(* CoDeSys 2.3 export: ld.exp *)

(* POU PLC_LD_PRG_TR, LD *)
PROGRAM PLC_LD_PRG_TR
VAR
END_VAR
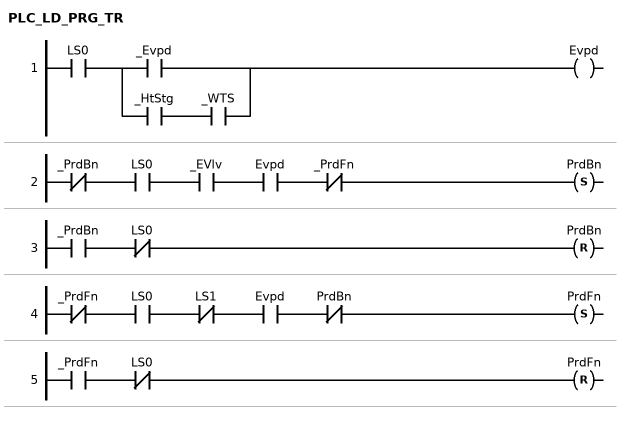
_LD_ (* Ladder Diagram *)
NETWORK 1
	[LS0] - { [_Evpd] | [_HtStg] - [_WTS] } --- (Evpd)
NETWORK 2
	[/_PrdBn] - [LS0] - [_EVlv] - [Evpd] - [/_PrdFn] --- (S PrdBn)
NETWORK 3
	[_PrdBn] - [/LS0] --- (R PrdBn)
NETWORK 4
	[/_PrdFn] - [LS0] - [/LS1] - [Evpd] - [/PrdBn] --- (S PrdFn)
NETWORK 5
	[_PrdFn] - [/LS0] --- (R PrdFn)
_END_LD_
(* the same logic as Structured Text *)
(* Network 1 *)
Evpd := LS0 AND (_Evpd OR _HtStg AND _WTS);
(* Network 2 *)
IF NOT _PrdBn AND LS0 AND _EVlv AND Evpd AND NOT _PrdFn THEN PrdBn := TRUE; END_IF;
(* Network 3 *)
IF _PrdBn AND NOT LS0 THEN PrdBn := FALSE; END_IF;
(* Network 4 *)
IF NOT _PrdFn AND LS0 AND NOT LS1 AND Evpd AND NOT PrdBn THEN PrdFn := TRUE; END_IF;
(* Network 5 *)
IF _PrdFn AND NOT LS0 THEN PrdFn := FALSE; END_IF;
END_PROGRAM
